ORGANIZATION_BLOCK "Main"
{ S7_Optimized_Access := 'TRUE' }
VERSION : 0.1
BEGIN
    "GDB_OperationsTest"();
    "FRK_TestPublish"(Complete := "GDB_OperationsTest".Done, Image0 := DWORD#2462965187, Image1 := DWORD#2239286705, Image2 := DWORD#1160051429, Image3 := DWORD#1259614334, Image4 := DWORD#648786163, Image5 := DWORD#284403629, Image6 := DWORD#210456493, Image7 := DWORD#4053867585, Result := "GDB_OperationsTest".Result, Status := "GDB_OperationsResultTest".Status);
END_ORGANIZATION_BLOCK
